FUNCTION_BLOCK T_ListOfNotificationHandlers
VAR_GENERIC CONSTANT
    MaxItems : UDINT := 10;
END_VAR
VAR
    _Count : UDINT;
    Items  : ARRAY[0..MaxItems - 1] OF I_NotificationHandler;
END_VAR

METHOD AddHandler
VAR_INPUT
    Handler : I_NotificationHandler;
END_VAR
IF _Count < MaxItems THEN
	Items[Count] := Handler;
	F_Inc(_Count);
END_IF
END_METHOD

METHOD Clear
VAR_INPUT
END_VAR
F_ClearMem(Items);
_Count := 0;
END_METHOD

PROPERTY Count : UDINT
GET
Count := _Count;
END_GET
END_PROPERTY

PROPERTY Full : BOOL
GET
Full := _Count >= MaxItems;
END_GET
END_PROPERTY

METHOD GetHandler : I_NotificationHandler
VAR_INPUT
    Index : UDINT;
END_VAR
IF Index < _Count THEN
    GetHandler := Items[Index];
END_IF
END_METHOD

METHOD HandlerInList : BOOL
VAR_INPUT
    HandlerToFind : I_NotificationHandler;
END_VAR
VAR
    NextHandler : I_NotificationHandler;
    i           : UDINT;
END_VAR
IF _Count < 1 THEN
    RETURN;
END_IF

FOR i := 0 TO _Count - 1 DO
    NextHandler := GetHandler(i);
    IF NextHandler = HandlerToFind THEN
        HandlerInList := TRUE;
    END_IF
END_FOR
END_METHOD

METHOD RemoveHandler
VAR_INPUT
    HandlerToRemove : I_NotificationHandler;
END_VAR
VAR
    NextHandler         : I_NotificationHandler;
    i                   : UDINT;
    RemovedHandlerIndex : UDINT;
    HandlerFound        : BOOL;
	LastHandlerIndex : UDINT;
END_VAR
IF _Count < 1 THEN
    RETURN;
END_IF

LastHandlerIndex := _Count - 1;

FOR i := 0 TO LastHandlerIndex DO
    // Get next handler...
    NextHandler := Items[i];

    // See if it the handler to remove...
    IF NextHandler = HandlerToRemove THEN
        RemovedHandlerIndex := i;
        HandlerFound        := TRUE;
    END_IF
END_FOR

IF HandlerFound THEN
    Items[RemovedHandlerIndex] := 0;

    IF RemovedHandlerIndex < LastHandlerIndex THEN
        // Shuffle remaining handlers...
		FOR i := RemovedHandlerIndex TO LastHandlerIndex - 1 DO
			Items[i] := Items[i + 1];
		END_FOR
		
    END_IF
    _Count := _Count - 1;

END_IF
END_METHOD

END_FUNCTION_BLOCK

(* stored: Version 1.1.0.1, ProductVersion 3.1.4026.19
   POU T_ListOfNotificationHandlers: Id {efdcf796-9d31-441b-a99c-4fd4a473f98e}, SpecialFunc None
   Folder Methods: Id {3d114acc-040e-4e27-8558-4e85fd10eea6}
   Folder Properties: Id {5d90d975-848f-4a9f-a35b-3776ce125fd4}
   Method AddHandler: Id {f0f02ca8-b2d4-4255-877a-514fb694031d}
   Method Clear: Id {b8dd6654-a37d-4b8a-bea5-3d7513a7295a}
   Property Count: Id {8898362c-5f01-4d65-b805-e83211742bad}
   Get Get: Id {8f67f0dd-fe96-4929-95fe-2afe73d0f3af}
   Property Full: Id {317243b2-18b4-47c6-aadd-b8ef5990c13f}
   Get Get: Id {4f799741-0f42-44e9-81a6-6b3c1b4f24b2}
   Method GetHandler: Id {86fce3f8-1332-44cb-87b7-dff84ff95854}
   Method HandlerInList: Id {23038192-9103-44af-a66f-062d5347818b}
   Method RemoveHandler: Id {41fc765e-18fa-4390-bc72-51ab9c6a726b} *)
